(* IEC 61131-3 sources: kns-port-domestic/tools/inventory_tests/fixtures/app/src/GVLs, 3 files *)

(* ---- GVL_Io.gvl.st ---- *)
// Сигналы ввода-вывода
VAR_GLOBAL
    xIn AT %I* : BOOL;
    xOut AT %QX0.1 : BOOL;
    wFlags AT %MW10 : WORD;
END_VAR

(* ---- GVL_Retain.gvl.st ---- *)
// Энергонезависимые переменные
VAR_GLOBAL RETAIN
    udiStarts : UDINT;
END_VAR
VAR_GLOBAL PERSISTENT RETAIN
    lrHours : LREAL;
END_VAR

(* ---- PersistentVars.pvl.st ---- *)
VAR_GLOBAL PERSISTENT RETAIN
    udiTrips : UDINT;
END_VAR
